Fanuc KAREL source: KA00227.KL

PROGRAM KA00227
%NOLOCKGROUP
VAR
  SRC: QUEUE_TYPE
  DST: QUEUE_TYPE
BEGIN
  DST = SRC
END KA00227
